(* IEC 61131-3 sources: MotionTestBenchMaster/Logical/30_MC/Libraries/MpAlarmX, 3 files *)

(* ---- MpAlarmX.typ ---- *)
(*Enumerations*)

TYPE
	MpAlarmXListUIStatusEnum :
		(
		mpALARMX_LIST_UI_STATUS_IDLE := 0, (*Indicates that no process is currently active*)
		mpALARMX_LIST_UI_STATUS_ERROR := 99 (*The last operation generated an error*)
		);
	MpAlarmXStateEnum :
		(
		mpALARMX_STATE_NONE := 0, (*Default state, alarm is not enabled*)
		mpALARMX_STATE_ACTIVE := 1, (*Active state, according OPC UA state model*)
		mpALARMX_STATE_INACTIVE := 2, (*Inactive state, according OPC UA state model*)
		mpALARMX_STATE_ACKNOWLEDGED := 3, (*Acknowledged state, according OPC UA state model*)
		mpALARMX_STATE_UNACKNOWLEDGED := 4 (*Unacknowledged state, according OPC UA state model*)
		);
	MpAlarmXAcknowledgeConfigEnum :
		(
		mpALARMX_ACK_DISABLED := 0, (*No acknowledgement required, inactive alarms disappear from current alarm list automatically.*)
		mpALARMX_ACK_REQ := 1, (*The alarm must be acknowledged, can be done at any time.*)
		mpALARMX_ACK_REQ_AFTER_ACTIVE := 2 (*The alarm must be acknowledged, can only be done when the alarm is inactive.*)
		);
	MpAlarmXHistoryUIStatusEnum :
		(
		mpALARMX_HISTORY_UI_STATUS_IDLE := 0, (*Indicates that no process is currently active*)
		mpALARMX_HISTORY_UI_STATUS_ERROR := 99 (*The last operation generated an error*)
		);
END_TYPE

(*FB Info Types*)

TYPE
	MpAlarmXStatusIDType : 	STRUCT
		ID : MpAlarmXErrorEnum; (*StatusID as enumerator*)
		Severity : MpComSeveritiesEnum; (*Severity of the error*)
		Code : UINT; (*Error code*)
	END_STRUCT;
	MpAlarmXDiagType : 	STRUCT
		StatusID : MpAlarmXStatusIDType; (*Segmented StatusID output*)
	END_STRUCT;
	MpAlarmXInfoType : 	STRUCT
		Diag : MpAlarmXDiagType; (*Additional diagnostic information*)
	END_STRUCT;
END_TYPE

(*UIConnect Types*)

TYPE
	MpAlarmXListUIBacktraceType : 	STRUCT
		RecordID : ARRAY[0..4]OF UDINT; (*The record ID of the logbook entry*)
		LogbookName : ARRAY[0..4]OF STRING[100]; (*The name of the logbook*)
		EventID : ARRAY[0..4]OF DINT; (*The event ID of the logbook entry*)
		Description : ARRAY[0..4]OF STRING[255]; (*The description text of this event ID*)
	END_STRUCT;
	MpAlarmXListUIAlarmListType : 	STRUCT
		Severity : ARRAY[0..49]OF UDINT; (*Alarm severity*)
		Code : ARRAY[0..49]OF UDINT; (*Alarm code*)
		Message : ARRAY[0..49]OF WSTRING[255]; (*Message describing the alarm*)
		AdditionalInformation1 : ARRAY[0..49]OF WSTRING[255]; (*A link with addidional information*)
		AdditionalInformation2 : ARRAY[0..49]OF WSTRING[255]; (*A link with addidional information*)
		InstanceID : ARRAY[0..49]OF UDINT; (*Unique alarm identity*)
		Scope : ARRAY[0..49]OF STRING[255]; (*The scope of the alarm*)
		Name : ARRAY[0..49]OF STRING[255]; (*Unique alarm name within the current scope*)
		StateActive : ARRAY[0..49]OF BOOL; (*Alarm is in Active state (according OPC UA Part 9: Alarms and Conditions)*)
		StateAcknowledged : ARRAY[0..49]OF BOOL; (*Alarm is in Acknowledged state (according OPC UA Part 9: Alarms and Conditions)*)
		Timestamp : ARRAY[0..49]OF STRING[50]; (*Timestamp of when the alarm was set*)
		SelectedIndex : UINT; (*The index of the currently selected alarm*)
		MaxSelection : UINT; (*The index of the last available alarm*)
		PageUp : BOOL; (*Command: Page Up (Scroll Up)*)
		PageDown : BOOL; (*Command: Page Down (Scroll Down)*)
		StepUp : BOOL; (*Command: Line Up (Scroll Up)*)
		StepDown : BOOL; (*Command: Line Down (Scroll Down)*)
		RangeStart : REAL; (*Displayed range: Start %*)
		RangeEnd : REAL; (*Displayed range: End %*)
	END_STRUCT;
	MpAlarmXListUIDetailsType : 	STRUCT
		Severity : UDINT; (*Alarm severity*)
		Code : UDINT; (*Alarm code*)
		Message : WSTRING[255]; (*Message describing the alarm*)
		AdditionalInformation1 : WSTRING[255]; (*A link with addidional information*)
		AdditionalInformation2 : WSTRING[255]; (*A link with addidional information*)
		InstanceID : UDINT; (*Unique alarm identity*)
		Scope : STRING[255]; (*The scope of the alarm*)
		Name : STRING[255]; (*Unique alarm name within the current scope*)
		StateActive : BOOL; (*Alarm is in Active state (according OPC UA Part 9: Alarms and Conditions)*)
		StateAcknowledged : BOOL; (*Alarm is in Acknowledged state (according OPC UA Part 9: Alarms and Conditions)*)
		Timestamp : STRING[50]; (*Timestamp of when the alarm was set*)
		Backtrace : MpAlarmXListUIBacktraceType; (*Backtrace of the alarm (origin logger entries)*)
	END_STRUCT;
	MpAlarmXListUIConnectType : 	STRUCT
		Status : MpAlarmXListUIStatusEnum; (*Current operation*)
		AlarmList : MpAlarmXListUIAlarmListType; (*List of available alarms*)
		Acknowledge : BOOL; (*Command: Acknowledge the selected alarm*)
		AcknowledgeAll : BOOL; (*Command: Acknowledge all alarms*)
		Details : MpAlarmXListUIDetailsType; (*Currently selected alarm*)
		Language : STRING[20]; (*Language ID that should be used when displaying data*)
		AcknowledgeID : UDINT; (*Command: Acknowledge the alarm with this instance ID*)
	END_STRUCT;
	MpAlarmXListUISetupType : 	STRUCT
		AlarmListSize : UINT := 20; (*Alarm list size*)
		AlarmListScrollWindow : USINT := 1; (*Scroll window (overlap for PageUp/Down)*)
		TimeStampPattern : STRING[50] := '%Y-%m-%d %H:%M:%S:%L'; (*Format pattern for the timestamp shown in the UIConnect structure. See MpAlarmXHistory configuration for details about the pattern syntax.*)
	END_STRUCT;
	MpAlarmXHistoryUIAlarmListType : 	STRUCT
		Severity : ARRAY[0..49]OF UDINT; (*Alarm severity*)
		Code : ARRAY[0..49]OF UDINT; (*Alarm code*)
		Message : ARRAY[0..49]OF WSTRING[255]; (*Message describing the alarm*)
		AdditionalInformation1 : ARRAY[0..49]OF WSTRING[255]; (*A link with addidional information*)
		AdditionalInformation2 : ARRAY[0..49]OF WSTRING[255]; (*A link with addidional information*)
		Scope : ARRAY[0..49]OF STRING[255]; (*The scope of the alarm*)
		Name : ARRAY[0..49]OF STRING[255]; (*Unique alarm name within the current scope*)
		OldState : ARRAY[0..49]OF MpAlarmXStateEnum; (*State change of this entry - the old state (according OPC UA Part 9: Alarms and Conditions)*)
		NewState : ARRAY[0..49]OF MpAlarmXStateEnum; (*State change of this entry - the new state (according OPC UA Part 9: Alarms and Conditions)*)
		Timestamp : ARRAY[0..49]OF STRING[50]; (*Timestamp of the state change (from OldState to NewState)*)
		SelectedIndex : UINT; (*The index of the currently selected alarm*)
		MaxSelection : UINT; (*The index of the last available alarm*)
		PageUp : BOOL; (*Command: Page Up (Scroll Up)*)
		PageDown : BOOL; (*Command: Page Down (Scroll Down)*)
		StepUp : BOOL; (*Command: Line Up (Scroll Up)*)
		StepDown : BOOL; (*Command: Line Down (Scroll Down)*)
		RangeStart : REAL; (*Displayed range: Start %*)
		RangeEnd : REAL; (*Displayed range: End %*)
	END_STRUCT;
	MpAlarmXHistoryUIDetailsType : 	STRUCT
		Severity : UDINT; (*Alarm severity*)
		Code : UDINT; (*Alarm code*)
		Message : WSTRING[255]; (*Message describing the alarm*)
		AdditionalInformation1 : WSTRING[255]; (*A link with addidional information*)
		AdditionalInformation2 : WSTRING[255]; (*A link with addidional information*)
		Scope : STRING[255]; (*The scope of the alarm*)
		Name : STRING[255]; (*Unique alarm name within the current scope*)
		OldState : MpAlarmXStateEnum; (*State change of this entry - the old state (according OPC UA Part 9: Alarms and Conditions)*)
		NewState : MpAlarmXStateEnum; (*State change of this entry - the new state (according OPC UA Part 9: Alarms and Conditions)*)
		Timestamp : STRING[50]; (*Timestamp of the state change (from OldState to NewState)*)
		DataDescriptions : ARRAY[0..9]OF STRING[50]; (*List of attached data to the alarm: data descriptions*)
		DataValues : ARRAY[0..9]OF STRING[255]; (*List of attached data to the alarm: data values*)
	END_STRUCT;
	MpAlarmXHistoryUIConnectType : 	STRUCT
		Status : MpAlarmXHistoryUIStatusEnum; (*Current operation*)
		AlarmList : MpAlarmXHistoryUIAlarmListType; (*List of available alarms*)
		Details : MpAlarmXHistoryUIDetailsType; (*Currently selected alarm*)
		Language : STRING[20]; (*Language ID that should be used when displaying data*)
	END_STRUCT;
	MpAlarmXHistoryUISetupType : 	STRUCT
		AlarmListSize : UINT := 20; (*Alarm list size*)
		AlarmListScrollWindow : USINT := 1; (*Scroll window (overlap for PageUp/Down)*)
		TimeStampPattern : STRING[50] := '%Y-%m-%d %H:%M:%S:%L'; (*Format pattern for the timestamp shown in the UIConnect structure. See MpAlarmXHistory configuration for details about the pattern syntax.*)
	END_STRUCT;
END_TYPE

(*Configuration Types*)

TYPE
	MpAlarmXMappingTypeEnum :
		(
		mpALARMX_MAPPING_TYPE_ALARM_NAME := 0, (*Load/Save a mapping by AlarmName from/to the configuration*)
		mpALARMX_MAPPING_TYPE_SEVERITY := 1, (*Load/Save a mapping by Severity from/to the configuration*)
		mpALARMX_MAPPING_TYPE_DEFAULT := 2 (*Load/Save a default mapping from/to the configuration*)
		);
	MpAlarmXActionEnum :
		(
		mpALARMX_ACT_NONE := 0, (*No action*)
		mpALARMX_ACT_REACTION := 1, (*Local reaction which can be evaluated with the MpAlarmXCheckReaction function*)
		mpALARMX_ACT_ESCALATE_ALARM := 2, (*Alarm is escalated by one level to the parent alarm core*)
		mpALARMX_ACT_ESCALATE_REACTION := 3, (*Reaction escalated by one level to the parent alarm core, can be evaluated with the MpAlarmXCheckReaction function there*)
		mpALARMX_ACT_REPLACE_ALARM := 4, (*Alarm is replaced by another alarm which is escalated by one level to the parent alarm core*)
		mpALARMX_ACT_SEND_MESSAGE := 5, (*Message is sent via MpTweet*)
		mpALARMX_ACT_REMAIN := 6 (*Alarm is remaining at this level*)
		);
	MpAlarmXActionConfigType : 	STRUCT  (*Defines configuration of one action*)
		Type : MpAlarmXActionEnum := 0; (*Reaction, Escalate, Replace, etc.*)
		Name : STRING[255] := ''; (*The meaning of this parameter depends on the Type, e.g. it is the alarm name for the ReplaceAlarm type, but the reaction name for the Reaction type*)
	END_STRUCT;
	MpAlarmXMappingConfigType : 	STRUCT  (*Configuration structure for the MpAlarmXConfigMapping FB*)
		Action : ARRAY[0..19]OF MpAlarmXActionConfigType; (*List of actions that should be performed with this mapping*)
	END_STRUCT;
	MpAlarmXAlarmConfigType : 	STRUCT  (*Configuration structure for the MpAlarmXConfigAlarm FB*)
		Message : STRING[255] := ''; (*The description text which the operator will see on the screen. Can include format items and references to the text system.*)
		Code : UDINT := 0; (*Numeric alarm code*)
		Severity : UDINT := 1; (*Severity is an indication of the urgency of an alarm, commonly also called Priority.*)
		Behavior : MpAlarmXBehaviorType; (*Select the pattern for the behavior options (Open advanced view for details: auto reset, auto acknowledge, recording options).*)
		Disable : BOOL := FALSE; (*The description text which the operator will see on the screen. Can include format items and references to the text system.*)
		AdditionalInformation1 : STRING[255] := ''; (*The description text which the operator will see on the screen. Can include format items and references to the text system.*)
		AdditionalInformation2 : STRING[255] := ''; (*The description text which the operator will see on the screen. Can include format items and references to the text system.*)
	END_STRUCT;
	MpAlarmXBehaviorType : 	STRUCT  (*Configuration structure of alarm behavior*)
		AutoReset : BOOL := FALSE; (*Alarm should be reset automatically immediately after being set (no subsequent call of MpAlarmXReset necessary).*)
		Acknowledge : MpAlarmXAcknowledgeConfigEnum := mpALARMX_ACK_REQ; (*Acknowledge behavior*)
		MultipleInstances : BOOL := FALSE; (*Multiple instances of this alarm should be possible.*)
		ReactionUntilAcknowledged : BOOL := TRUE; (*Any reactions caused by the alarm will remain active until the alarm is acknowledged.*)
		HistoryReport : MpAlarmXHistoryReportType; (*Define which state changes should be recorded for historical logging.*)
	END_STRUCT;
	MpAlarmXHistoryReportType : 	STRUCT  (*Define which state changes should be recorded for historical logging.*)
		InactiveToActive : BOOL := TRUE; (*State changes from Inactive to Active should be recorded.*)
		ActiveToInactive : BOOL := TRUE; (*State changes from Active to Inactive should be recorded.*)
		UnacknowledgedToAcknowledged : BOOL := TRUE; (*State changes from Unacknowledged to Acknowledged should be recorded.*)
	END_STRUCT;
END_TYPE

(* ---- MpAlarmXError.typ ---- *)
TYPE
    MpAlarmXErrorEnum :
        ( (* Error numbers of library MpAlarmX *)
        mpALARMX_NO_ERROR := 0, (* No error *)
        mpALARMX_ERR_ACTIVATION := -1064239103, (* Could not create component [Error: 1, 0xc0910001] *)
        mpALARMX_ERR_MPLINK_NULL := -1064239102, (* MpLink is NULL pointer [Error: 2, 0xc0910002] *)
        mpALARMX_ERR_MPLINK_INVALID := -1064239101, (* MpLink connection not allowed [Error: 3, 0xc0910003] *)
        mpALARMX_ERR_MPLINK_CHANGED := -1064239100, (* MpLink modified [Error: 4, 0xc0910004] *)
        mpALARMX_ERR_MPLINK_CORRUPT := -1064239099, (* Invalid MpLink contents [Error: 5, 0xc0910005] *)
        mpALARMX_ERR_MPLINK_IN_USE := -1064239098, (* MpLink already in use [Error: 6, 0xc0910006] *)
        mpALARMX_ERR_CONFIG_NULL := -1064239096, (* Configuration structure is null pointer [Error: 8, 0xc0910008] *)
        mpALARMX_ERR_CONFIG_INVALID := -1064239091, (* Invalid Configuration [Error: 13, 0xc091000d] *)
        mpALARMX_ERR_NAME_NULL := -1064116224, (* The specified name is NULL [Error: 57344, 0xc092e000] *)
        mpALARMX_ERR_NAME_EMPTY := -1064116223, (* The specified name is empty [Error: 57345, 0xc092e001] *)
        mpALARMX_WRN_MISSING_UICONNECT := -2137858045, (* UIConnect is NULL [Warning: 57347, 0x8092e003] *)
        mpALARMX_ERR_ALARM_NOT_ACTIVE := -1064116220, (* The alarm is unknown and cannot be reset [Error: 57348, 0xc092e004] *)
        mpALARMX_ERR_ALARM_NOT_SELECTED := -1064116219, (* No alarm is selected [Error: 57349, 0xc092e005] *)
        mpALARMX_ERR_ACK_NOT_ALLOWED := -1064116218, (* The alarm cannot be acknowledged at this position in the component tree [Error: 57350, 0xc092e006] *)
        mpALARMX_ERR_INVALID_FILE_DEV := -1064116217, (* The specified device name in NULL [Error: 57351, 0xc092e007] *)
        mpALARMX_INF_WAIT_CORE_FB := 1083367432, (* Waiting for parent component [Informational: 57352, 0x4092e008] *)
        mpALARMX_ERR_CORE_INST_EXISTS := -1064116215, (* Another core component was already found in this component group [Error: 57353, 0xc092e009] *)
        mpALARMX_ERR_MEMORY_INIT := -1064116214, (* The history memory could not be initialized. See log for furher details [Error: 57354, 0xc092e00a] *)
        mpALARMX_ERR_WRITE_EXPORT_FILE := -1064116213, (* Error while writing to the history export file [Error: 57355, 0xc092e00b] *)
        mpALARMX_ERR_NAME_NOT_FOUND := -1064116212 (* The specified alarm name was not found [Error: 57356, 0xc092e00c] *)
        );
END_TYPE

(* ---- MpAlarmX.fun ---- *)
(*Core Function Blocks*)

FUNCTION_BLOCK MpAlarmXCore (*mapp component for advanced centralized alarm collection and management*) (* $GROUP=mapp,$CAT=Alarm System,$GROUPICON=Icon_mapp.png,$CATICON=Icon_MpAlarmX.png *)
	VAR_INPUT
		MpLink : REFERENCE TO MpComIdentType; (*Incoming communication handle (mapp standard interface)*) (* *) (*#PAR#;*)
		Enable : BOOL; (*Enables/Disables the function block (mapp standard interface)*) (* *) (*#PAR#;*)
		ErrorReset : BOOL; (*Resets all function block errors (mapp standard interface)*) (* *) (*#PAR#;*)
	END_VAR
	VAR_OUTPUT
		Active : BOOL; (*Function block is active (mapp standard interface)*) (* *) (*#PAR#;*)
		Error : BOOL; (*Indicates an error (mapp standard interface)*) (* *) (*#PAR#;*)
		StatusID : DINT; (*Error/Status information (mapp standard interface)*) (* *) (*#PAR#; *)
		ActiveAlarms : UDINT; (*Number of alarms which are currently active*) (* *) (*#CMD#;*)
		PendingAlarms : UDINT; (*Number of alarms which are currently pending (either active, or not yet acknowleged)*) (* *) (*#CMD#;*)
		Info : MpAlarmXInfoType; (*Additional information*) (* *) (*#CMD#;*)
	END_VAR
	VAR
		Internal : {REDUND_UNREPLICABLE} MpComInternalDataType; (*Internal data*) (* *) (*#OMIT#;*)
	END_VAR
END_FUNCTION_BLOCK
(*UI Function Blocks*)

FUNCTION_BLOCK MpAlarmXListUI (*add-on function block that provides VC4 connection datapoints to display the currently active alarms in a list*) (* $GROUP=mapp,$CAT=Alarm System,$GROUPICON=Icon_mapp.png,$CATICON=Icon_MpAlarmX.png *)
	VAR_INPUT
		MpLink : REFERENCE TO MpComIdentType; (*Incoming communication handle (mapp standard interface)*) (* *) (*#PAR#;*)
		Enable : BOOL; (*Enables/Disables the function block (mapp standard interface)*) (* *) (*#PAR#;*)
		ErrorReset : BOOL; (*Resets all function block errors (mapp standard interface)*) (* *) (*#PAR#;*)
		UISetup : MpAlarmXListUISetupType; (*Setup UI connection - must be configured before enabling the FB*) (* *) (*#PAR#;*)
		UIConnect : REFERENCE TO MpAlarmXListUIConnectType; (*UI connection datapoints*) (* *) (*#CMD#;*)
	END_VAR
	VAR_OUTPUT
		Active : BOOL; (*Function block is active (mapp standard interface)*) (* *) (*#PAR#;*)
		Error : BOOL; (*Indicates an error (mapp standard interface)*) (* *) (*#PAR#;*)
		StatusID : DINT; (*Error/Status information (mapp standard interface)*) (* *) (*#PAR#; *)
		Info : MpAlarmXInfoType; (*Additional information*) (* *) (*#CMD#;*)
	END_VAR
	VAR
		Internal : {REDUND_UNREPLICABLE} MpComInternalDataType; (*Internal data*) (* *) (*#OMIT#;*)
	END_VAR
END_FUNCTION_BLOCK

FUNCTION_BLOCK MpAlarmXHistoryUI (*add-on function block that provides VC4 connection datapoints to display the alarm history in a list*) (* $GROUP=mapp,$CAT=Alarm System,$GROUPICON=Icon_mapp.png,$CATICON=Icon_MpAlarmX.png *)
	VAR_INPUT
		MpLink : REFERENCE TO MpComIdentType; (*Incoming communication handle (mapp standard interface)*) (* *) (*#PAR#;*)
		Enable : BOOL; (*Enables/Disables the function block (mapp standard interface)*) (* *) (*#PAR#;*)
		ErrorReset : BOOL; (*Resets all function block errors (mapp standard interface)*) (* *) (*#PAR#;*)
		UISetup : MpAlarmXHistoryUISetupType; (*Setup UI connection - must be configured before enabling the FB*) (* *) (*#PAR#;*)
		UIConnect : REFERENCE TO MpAlarmXHistoryUIConnectType; (*UI connection datapoints*) (* *) (*#CMD#;*)
	END_VAR
	VAR_OUTPUT
		Active : BOOL; (*Function block is active (mapp standard interface)*) (* *) (*#PAR#;*)
		Error : BOOL; (*Indicates an error (mapp standard interface)*) (* *) (*#PAR#;*)
		StatusID : DINT; (*Error/Status information (mapp standard interface)*) (* *) (*#PAR#; *)
		Info : MpAlarmXInfoType; (*Additional information*) (* *) (*#CMD#;*)
	END_VAR
	VAR
		Internal : {REDUND_UNREPLICABLE} MpComInternalDataType; (*Internal data*) (* *) (*#OMIT#;*)
	END_VAR
END_FUNCTION_BLOCK
(*General add-ons*)

FUNCTION MpAlarmXCheckState : BOOL (*Add-on function which checks whether an alarm is currently in a certain state*) (* $GROUP=mapp,$CAT=Alarm System,$GROUPICON=Icon_mapp.png,$CATICON=Icon_MpAlarmX.png *)
	VAR_INPUT
		MpLink : MpComIdentType; (*Incoming communication handle (mapp standard interface)*) (* *) (*#PAR#;*)
		Name : STRING[255]; (*Unique Identifier of the alarm*) (* *) (*#PAR#;*)
		State : MpAlarmXStateEnum; (*Check whether the alarm is currently in this state*) (* *) (*#PAR#;*)
	END_VAR
END_FUNCTION

FUNCTION MpAlarmXCheckStateID : BOOL (*Add-on function which checks whether an alarm is currently in a certain state*) (* $GROUP=mapp,$CAT=Alarm System,$GROUPICON=Icon_mapp.png,$CATICON=Icon_MpAlarmX.png *)
	VAR_INPUT
		MpLink : MpComIdentType; (*Incoming communication handle (mapp standard interface)*) (* *) (*#PAR#;*)
		InstanceID : UDINT; (*Instance ID of the alarm that should be checked for its state*) (* *) (*#PAR#;*)
		State : MpAlarmXStateEnum; (*Check whether the alarm is currently in this state*) (* *) (*#PAR#;*)
	END_VAR
END_FUNCTION

FUNCTION MpAlarmXCheckReaction : BOOL (*Add-on function which checks whether a certain reaction is currently active, returns TRUE if at least one alarm is currently active that requires this reaction*) (* $GROUP=mapp,$CAT=Alarm System,$GROUPICON=Icon_mapp.png,$CATICON=Icon_MpAlarmX.png *)
	VAR_INPUT
		MpLink : MpComIdentType; (*Incoming communication handle (mapp standard interface)*) (* *) (*#PAR#;*)
		Name : STRING[255]; (*Unique name of the reaction*) (* *) (*#PAR#;*)
	END_VAR
END_FUNCTION

FUNCTION MpAlarmXSet : UDINT (*Add-On function to set (raise) a user alarm. By calling this function the alarm system is informed that a specific alarm is active. Returns InstanceID of the alarm that was set.*) (* $GROUP=mapp,$CAT=Alarm System,$GROUPICON=Icon_mapp.png,$CATICON=Icon_MpAlarmX.png *)
	VAR_INPUT
		MpLink : MpComIdentType; (*Incoming communication handle (mapp standard interface)*) (* *) (*#PAR#;*)
		Name : STRING[255]; (*Unique name of the alarm*) (* *) (*#PAR#;*)
	END_VAR
END_FUNCTION

FUNCTION MpAlarmXAcknowledge : DINT (*Add-On function to acknowledge an alarm. By calling this function the alarm system is informed that the operator has acknowledged an alarm. Returns result code.*) (* $GROUP=mapp,$CAT=Alarm System,$GROUPICON=Icon_mapp.png,$CATICON=Icon_MpAlarmX.png *)
	VAR_INPUT
		MpLink : MpComIdentType; (*Incoming communication handle (mapp standard interface)*) (* *) (*#PAR#;*)
		Name : STRING[255]; (*Unique name of the alarm*) (* *) (*#PAR#;*)
	END_VAR
END_FUNCTION

FUNCTION MpAlarmXAcknowledgeID : DINT (*Add-On function to acknowledge an alarm. By calling this function the alarm system is informed that the operator has acknowledged an alarm. Returns result code.*) (* $GROUP=mapp,$CAT=Alarm System,$GROUPICON=Icon_mapp.png,$CATICON=Icon_MpAlarmX.png *)
	VAR_INPUT
		MpLink : MpComIdentType; (*Incoming communication handle (mapp standard interface)*) (* *) (*#PAR#;*)
		InstanceID : UDINT; (*Instance ID of the alarm that should be acknowledged*) (* *) (*#PAR#;*)
	END_VAR
END_FUNCTION

FUNCTION MpAlarmXReset : DINT (*Add-On function to reset a user alarm. By calling this function the alarm system is informed that a specific alarm is inactive. Returns result code.*) (* $GROUP=mapp,$CAT=Alarm System,$GROUPICON=Icon_mapp.png,$CATICON=Icon_MpAlarmX.png *)
	VAR_INPUT
		MpLink : MpComIdentType; (*Incoming communication handle (mapp standard interface)*) (* *) (*#PAR#;*)
		Name : STRING[255]; (*Unique name of the alarm*) (* *) (*#PAR#;*)
	END_VAR
END_FUNCTION

FUNCTION MpAlarmXResetID : DINT (*Add-On function to reset a user alarm. By calling this function the alarm system is informed that a specific alarm is inactive. Returns result code.*) (* $GROUP=mapp,$CAT=Alarm System,$GROUPICON=Icon_mapp.png,$CATICON=Icon_MpAlarmX.png *)
	VAR_INPUT
		MpLink : MpComIdentType; (*Incoming communication handle (mapp standard interface)*) (* *) (*#PAR#;*)
		InstanceID : UDINT; (*Instance ID of the alarm that should be reset*) (* *) (*#PAR#;*)
	END_VAR
END_FUNCTION
(*History add-ons*)

FUNCTION_BLOCK MpAlarmXHistory (*Historical recording of all alarm related events*) (* $GROUP=mapp,$CAT=Alarm System,$GROUPICON=Icon_mapp.png,$CATICON=Icon_MpAlarmX.png *)
	VAR_INPUT
		MpLink : REFERENCE TO MpComIdentType; (*Incoming communication handle (mapp standard interface)*) (* *) (*#PAR#;*)
		Enable : BOOL; (*Enables/Disables the function block (mapp standard interface)*) (* *) (*#PAR#;*)
		ErrorReset : BOOL; (*Resets all function block errors (mapp standard interface)*) (* *) (*#PAR#;*)
		DeviceName : REFERENCE TO STRING[50]; (*Name of device to export the alarm history to*) (* *) (*#CMD#;*)
		Language : REFERENCE TO STRING[20]; (*Language ID that should be used when exporting data*) (* *) (*#CMD#OPT#;*)
		Export : BOOL; (*Save the current alarm history data (since last archiving) to the given file device (as a human-readable file)*) (* *) (*#CMD#;*)
	END_VAR
	VAR_OUTPUT
		Active : BOOL; (*Function block is active (mapp standard interface)*) (* *) (*#PAR#;*)
		Error : BOOL; (*Indicates an error (mapp standard interface)*) (* *) (*#PAR#;*)
		StatusID : DINT; (*Error/Status information (mapp standard interface)*) (* *) (*#PAR#; *)
		CommandBusy : BOOL; (*Function block is busy processing a command.*) (* *) (*#CMD#OPT#;*)
		CommandDone : BOOL; (*Command has finished and was successful.*) (* *) (*#CMD#;*)
		Info : MpAlarmXInfoType; (*Additional information*) (* *) (*#CMD#;*)
	END_VAR
	VAR
		Internal : {REDUND_UNREPLICABLE} MpComInternalDataType;
	END_VAR
END_FUNCTION_BLOCK
(*Configuration add-ons*)

FUNCTION_BLOCK MpAlarmXConfigAlarm (*add-on function block that allows to load and save alarm configurations *) (* $GROUP=mapp,$CAT=Alarm System,$GROUPICON=Icon_mapp.png,$CATICON=Icon_MpAlarmX.png *)
	VAR_INPUT
		MpLink : REFERENCE TO MpComIdentType; (*Incoming communication handle (mapp standard interface)*) (* *) (*#PAR#;*)
		Enable : BOOL; (*Enables/Disables the function block (mapp standard interface)*) (* *) (*#PAR#;*)
		ErrorReset : BOOL; (*Resets all function block errors (mapp standard interface)*) (* *) (*#PAR#;*)
		Name : REFERENCE TO STRING[255]; (*Unique Identifier of the alarm*) (* *) (*#PAR#;*)
		Configuration : REFERENCE TO MpAlarmXAlarmConfigType; (*Configuration parameters (mapp standard interface)*) (* *) (*#PAR#;*)
		Load : BOOL; (*Read configuration from AR into the config structure*) (* *) (*#CMD#*)
		Save : BOOL; (*Write configuration from config structure to AR*) (* *) (*#CMD#*)
	END_VAR
	VAR_OUTPUT
		Active : BOOL; (*Function block is active (mapp standard interface)*) (* *) (*#PAR#;*)
		Error : BOOL; (*Indicates an error (mapp standard interface)*) (* *) (*#PAR#;*)
		StatusID : DINT; (*Error/Status information (mapp standard interface)*) (* *) (*#PAR#; *)
		CommandBusy : BOOL; (*Function block is busy processing a command.*) (* *) (*#CMD#OPT#;*)
		CommandDone : BOOL; (*Command has finished and was successful.*) (* *) (*#CMD#*)
		Info : MpAlarmXInfoType; (*Additional information*) (* *) (*#CMD#;*)
	END_VAR
	VAR
		Internal : {REDUND_UNREPLICABLE} MpComInternalDataType; (*Internal data*)
	END_VAR
END_FUNCTION_BLOCK

FUNCTION_BLOCK MpAlarmXConfigMapping (*add-on function block that allows to load and save mapping configurations *) (* $GROUP=mapp,$CAT=Alarm System,$GROUPICON=Icon_mapp.png,$CATICON=Icon_MpAlarmX.png *)
	VAR_INPUT
		MpLink : REFERENCE TO MpComIdentType; (*Incoming communication handle (mapp standard interface)*) (* *) (*#PAR#;*)
		Enable : BOOL; (*Enables/Disables the function block (mapp standard interface)*) (* *) (*#PAR#;*)
		ErrorReset : BOOL; (*Resets all function block errors (mapp standard interface)*) (* *) (*#PAR#;*)
		Type : MpAlarmXMappingTypeEnum; (*Type of the mapping (Alarm Name, Severity or Default)*) (* *) (*#PAR#;*)
		Name : REFERENCE TO STRING[255]; (*Name (meaning depends on the Type setting)*) (* *) (*#PAR#;*)
		Configuration : REFERENCE TO MpAlarmXMappingConfigType; (*Configuration parameters (mapp standard interface)*) (* *) (*#PAR#;*)
		Load : BOOL; (*Read configuration from AR into the config structure*) (* *) (*#CMD#*)
		Save : BOOL; (*Write configuration from config structure to AR*) (* *) (*#CMD#*)
	END_VAR
	VAR_OUTPUT
		Active : BOOL; (*Function block is active (mapp standard interface)*) (* *) (*#PAR#;*)
		Error : BOOL; (*Indicates an error (mapp standard interface)*) (* *) (*#PAR#;*)
		StatusID : DINT; (*Error/Status information (mapp standard interface)*) (* *) (*#PAR#; *)
		CommandBusy : BOOL; (*Function block is busy processing a command.*) (* *) (*#CMD#OPT#;*)
		CommandDone : BOOL; (*Command has finished and was successful.*) (* *) (*#CMD#*)
		Info : MpAlarmXInfoType; (*Additional information*) (* *) (*#CMD#;*)
	END_VAR
	VAR
		Internal : {REDUND_UNREPLICABLE} MpComInternalDataType; (*Internal data*)
	END_VAR
END_FUNCTION_BLOCK
